(* PLC project Motor_StartStop_TM241CE24T, PLCAutoPilot M241 Generator 2.0 *)
(* stored: creationDateTime 2025-12-30T01:30:00, modificationDateTime 2025-12-30T01:30:00 *)

FUNCTION_BLOCK GVL_IO
  VAR
    StartPB : BOOL;  (* Start Pushbutton (NO) - Map to %IX0.0 *)
    StopPB : BOOL;  (* Stop Pushbutton (NC) - Map to %IX0.1 *)
    OverloadTrip : BOOL;  (* Thermal Overload (NC) - Map to %IX0.2 *)
    EmergencyStop : BOOL;  (* E-Stop (NC) - Map to %IX0.3 *)
    MotorContactor : BOOL;  (* Main Contactor - Map to %QX0.0 *)
    RunIndicator : BOOL;  (* Run Lamp - Map to %QX0.1 *)
    FaultIndicator : BOOL;  (* Fault Lamp - Map to %QX0.2 *)
  END_VAR

            
// GVL_IO - Global Variable List for Motor Start/Stop
// Map these variables to physical I/O addresses after import
            
          
END_FUNCTION_BLOCK

(* Motor Start/Stop Control Program (Structured Text) Features: - 3 second startup delay (anti-chatter) - Overload fault latching with automatic reset - Emergency stop interlock - Run and fault indication lamps Safety: - StopPB is NC (fail-safe: wire break = motor stops) - EmergencyStop is NC (fail-safe) - OverloadTrip is NC (fail-safe) Generated by PLCAutoPilot for TM241CE24T *)
PROGRAM Motor_Control_ST
  VAR
    MotorRunning : BOOL;  (* Motor Running Status *)
    MotorFault : BOOL;  (* Motor Fault Latched *)
    SafetyOK : BOOL;  (* Safety Interlock OK *)
    StartupTimer : TON;  (* 3 second startup delay *)
    IO : GVL_IO;  (* I/O Interface *)
  END_VAR

            
// ============================================
// MOTOR START/STOP CONTROL (Structured Text)
// TM241CE24T - PLCAutoPilot Generated
// ============================================
//
// I/O MAPPING (configure in GVL_IO instance):
// Inputs:
//   IO.StartPB       - %IX0.0 (NO pushbutton)
//   IO.StopPB        - %IX0.1 (NC pushbutton)
//   IO.OverloadTrip  - %IX0.2 (NC thermal relay)
//   IO.EmergencyStop - %IX0.3 (NC E-Stop)
//
// Outputs:
//   IO.MotorContactor - %QX0.0 (Main contactor K1)
//   IO.RunIndicator   - %QX0.1 (Run lamp)
//   IO.FaultIndicator - %QX0.2 (Fault lamp)
// ============================================

// Safety interlock check
// E-Stop must be OK (NC contact = TRUE when OK)
// Overload must be OK (NC contact = FALSE when OK)
SafetyOK := IO.EmergencyStop AND NOT IO.OverloadTrip;

// Fault latching
// Set fault when overload trips
IF IO.OverloadTrip THEN
    MotorFault := TRUE;
END_IF;

// Reset fault when Start is pressed AND overload is cleared
IF IO.StartPB AND NOT IO.OverloadTrip THEN
    MotorFault := FALSE;
END_IF;

// Startup timer (3 second anti-chatter delay)
// Timer runs when Start pressed, Safety OK, and no fault
StartupTimer(
    IN := IO.StartPB AND SafetyOK AND NOT MotorFault AND NOT MotorRunning,
    PT := T#3S
);

// Motor running logic
// SET: Timer complete (3 seconds of continuous Start press)
IF StartupTimer.Q THEN
    MotorRunning := TRUE;
END_IF;

// RESET: Stop pressed OR Safety NOT OK OR Fault
// Note: StopPB is NC, so FALSE = pressed
IF NOT IO.StopPB OR NOT SafetyOK OR MotorFault THEN
    MotorRunning := FALSE;
END_IF;

// Write to outputs
IO.MotorContactor := MotorRunning;
IO.RunIndicator := MotorRunning;
IO.FaultIndicator := MotorFault;
            
          
END_PROGRAM

(* Motor Start/Stop Control (Instruction List / Ladder equivalent) This program implements the same logic as Motor_Control_ST using Instruction List language which maps directly to Ladder rungs. Generated by PLCAutoPilot for TM241CE24T *)
PROGRAM Motor_Control_IL
  VAR
    MotorRunning : BOOL;
    MotorFault : BOOL;
    SafetyOK : BOOL;
    StartCondition : BOOL;
    StopCondition : BOOL;
    StartupTimer : TON;
    StartupComplete : BOOL;
    IO : GVL_IO;
  END_VAR

            
(* ============================================
   MOTOR START/STOP CONTROL (Instruction List)
   Equivalent to Ladder Diagram
   TM241CE24T - PLCAutoPilot Generated
   ============================================ *)

(* RUNG 1: Safety Interlock *)
LD    IO.EmergencyStop
ANDN  IO.OverloadTrip
ST    SafetyOK

(* RUNG 2: Fault Latch SET *)
LD    IO.OverloadTrip
S     MotorFault

(* RUNG 3: Fault Latch RESET *)
LD    IO.StartPB
ANDN  IO.OverloadTrip
R     MotorFault

(* RUNG 4: Start Conditions *)
LD    IO.StartPB
AND   SafetyOK
ANDN  MotorFault
ANDN  MotorRunning
ST    StartCondition

(* RUNG 5: Startup Timer *)
CAL   StartupTimer(IN := StartCondition, PT := T#3S)
LD    StartupTimer.Q
ST    StartupComplete

(* RUNG 6: Motor Latch SET *)
LD    StartupComplete
S     MotorRunning

(* RUNG 7: Stop Conditions *)
LDN   IO.StopPB
ORN   SafetyOK
OR    MotorFault
ST    StopCondition

(* RUNG 8: Motor Latch RESET *)
LD    StopCondition
R     MotorRunning

(* RUNG 9-11: Outputs *)
LD    MotorRunning
ST    IO.MotorContactor
ST    IO.RunIndicator
LD    MotorFault
ST    IO.FaultIndicator
            
          
END_PROGRAM

CONFIGURATION TM241CE24T
  RESOURCE Application ON PLC
    TASK MAST(INTERVAL := T#20ms, PRIORITY := 1);
    PROGRAM Motor_Control_ST_Inst WITH MAST : Motor_Control_ST;
  END_RESOURCE
END_CONFIGURATION
